Staubli VAL3: editIF.pgx

public program editIF(string x_sKey, num x_nIndex, string& x_sType[], string& x_sIOIndex[], num& x_nValue[], string x_sANDOR1, string x_sANDOR2, bool& x_bToSave)
  local num l_i
  local num l_nIndex
  local bool l_bResult
begin
  if x_nIndex==0 and progTemp:pProgItem[x_sKey].pProgTemplate[x_nIndex].sTRAJname==""
    x_nIndex=x_nIndex
  else
    x_nIndex=x_nIndex+1
    append(progTemp:pProgItem[x_sKey].pProgTemplate)
    for l_i = size(progTemp:pProgItem[x_sKey].pProgTemplate)-1 to x_nIndex step -1
      call copyPara(x_sKey,l_i-1,l_i)
    endFor
    //insert(progTemp:pProgItem[x_sKey].pProgTemplate[x_nIndex])
  endIf

  progTemp:pProgItem[x_sKey].pProgTemplate[x_nIndex].nType=3
  progTemp:pProgItem[x_sKey].pProgTemplate[x_nIndex].sTRAJname="IF"
  for l_i = 0 to 2
    if x_sIOIndex[l_i]!=""
      toNum(x_sIOIndex[l_i],l_nIndex,l_bResult)
    else
      l_nIndex=-1
    endIf
    switch x_sType[l_i]
      case "DIN"
        progTemp:pProgItem[x_sKey].pProgTemplate[x_nIndex].iIfItem.nSigType[l_i]=1
        progTemp:pProgItem[x_sKey].pProgTemplate[x_nIndex].iIfItem.nSigIndex[l_i]=l_nIndex
        progTemp:pProgItem[x_sKey].pProgTemplate[x_nIndex].iIfItem.nValue[l_i]=x_nValue[l_i]
      break
      case "DOUT"
        progTemp:pProgItem[x_sKey].pProgTemplate[x_nIndex].iIfItem.nSigType[l_i]=2
        progTemp:pProgItem[x_sKey].pProgTemplate[x_nIndex].iIfItem.nSigIndex[l_i]=l_nIndex
        progTemp:pProgItem[x_sKey].pProgTemplate[x_nIndex].iIfItem.nValue[l_i]=x_nValue[l_i]

      break
      case "AIN"
        progTemp:pProgItem[x_sKey].pProgTemplate[x_nIndex].iIfItem.nSigType[l_i]=3
        progTemp:pProgItem[x_sKey].pProgTemplate[x_nIndex].iIfItem.nSigIndex[l_i]=l_nIndex
        progTemp:pProgItem[x_sKey].pProgTemplate[x_nIndex].iIfItem.nValue[l_i]=x_nValue[l_i]

      break
      case "AOUT"
        progTemp:pProgItem[x_sKey].pProgTemplate[x_nIndex].iIfItem.nSigType[l_i]=4
        progTemp:pProgItem[x_sKey].pProgTemplate[x_nIndex].iIfItem.nSigIndex[l_i]=l_nIndex
        progTemp:pProgItem[x_sKey].pProgTemplate[x_nIndex].iIfItem.nValue[l_i]=x_nValue[l_i]

      break
      default
        progTemp:pProgItem[x_sKey].pProgTemplate[x_nIndex].iIfItem.nSigType[l_i]=0
        progTemp:pProgItem[x_sKey].pProgTemplate[x_nIndex].iIfItem.nSigIndex[l_i]=-1
        progTemp:pProgItem[x_sKey].pProgTemplate[x_nIndex].iIfItem.nValue[l_i]=0

      break
    endSwitch
  endFor

  progTemp:pProgItem[x_sKey].pProgTemplate[x_nIndex].iIfItem.bANDOR[0]=(x_sANDOR1=="OR")
  progTemp:pProgItem[x_sKey].pProgTemplate[x_nIndex].iIfItem.bANDOR[1]=(x_sANDOR2=="OR")

  x_bToSave=true
end
